Universal Robots PolyScope program: Sub_Centrifuge_V3.urp

Program Sub_Centrifuge_V3 (installation=default directory=/programs/03 Sub Routines createdIn=5.13.0 lastSavedIn=5.16.0 robotSerialNumber=20245590049)
Calibrated DH parameters: a=[0.000139, -0.197451, -0.383992, -0.000109, 0.000038, 0]; d=[0.162494, 274.063354, -251.846761, -22.083037, 0.099612, 0.099364]; alpha=[1.570089, 0.001374, 0.003592, 1.570222, -1.570187, 0]; deltaTheta=[0, 1.08787, 5.400214, -0.204909, 0.000001, 0]
InitVariablesNode variables(variable(name=DEV_CEN_PosRtr, expression=0))
BeforeStart
  Centrifuge := rpc_factory("xmlrpc","http://192.168.12.125:50002")
  Action :=  (valueSource=Operator message=What to do? valueType=Integer)
Robot Program (runOnlyOnce=true)
  Folder Handling
    SuppressedNode
      Folder PreSettings
        Folder Init Move Definitions [hidden by the author, left out]
        Folder Jig Definition [hidden by the author, left out]
        Folder Frame Definition [hidden by the author, left out]
        Folder Pose Definition [hidden by the author, left out]
    '===================='
    Switch expression=Action
      Case (caseValue=5)
        Folder Open
          Script: Centrifuge.open_hatch()
      Case (caseValue=6)
        Folder Close
          Script: Centrifuge.close_hatch()
      Case (caseValue=7)
        Folder Load
          DEV_CEN_CmdRslt := Centrifuge.move_rotor(DEV_CEN_PosRtr)
          If JNT_S≠[0,0,0,0,0,0]
            MoveJ speed 90 deg/s, acceleration 80 deg/s^2 (useActiveTCP=true positionType=JointAngles) feature=Base
              Waypoint Variable (Variable): motionParameters(blendRadius=0.05); variable=JNT_S
          MoveJ speed 90 deg/s, acceleration 80 deg/s^2 (useActiveTCP=true) feature=FRM_Reference
            If PSE_A_H≠p[0,0,0,0,0,0]
              Waypoint Variable (Variable): motionParameters(blendRadius=0.02); variable=PSE_A_H
            Waypoint Variable (Variable): variable=PSE_A
          If Centrifuge.posreached(DEV_CEN_PosRtr)
            MoveL speed 300 mm/s, acceleration 1200 mm/s^2 (useActiveTCP=true) feature=FRM_Reference
              If PSE_T_H≠p[0,0,0,0,0,0]
                Waypoint Variable (Variable): variable=PSE_T_H
              Waypoint Variable (Variable): motionParameters(jointSpeed=1.047198 jointAcceleration=1.396263 cartesianSpeed=0.075 cartesianAcceleration=1.2); variable=PSE_T
                Until TOOL_CONTACT_DETECTION (allowActions=true retraction=0.001 decelerationAcceleration=0.5 decelerationAngularAcceleration=34.906585)
                  Folder EOAT
                    URCap Gripper (Robotiq_Grippers, Robotiq Inc.) dataModel(position=88.72549019607843, force=25.0, speed=50.0, positionInDouble=88.72549019607843, forceInDouble=25.0, speedInDouble=50.0, slaveIds=[9], blocking=true)
                  Force Frame feature=Joint_6_name; selection=[0, 0, 0, 0, 0, 1]; wrench=[0, 0, 0, 0, 0, 0]; limitsForce=[0.15, 0.15, 0.15, 1.047198, 1.047198, 3.141593]; limitsMotion=[0.1, 0.1, 0.1, 0.349066, 0.349066, 0.349066]
                    Waypoint Variable (Variable): motionParameters(jointSpeed=1.047198 jointAcceleration=1.396263 cartesianSpeed=0.01 cartesianAcceleration=1.2); variable=PSE_T
              Folder EOAT
                URCap Gripper (Robotiq_Grippers, Robotiq Inc.) dataModel(position=70.09803921568627, force=50.0, speed=50.0, positionInDouble=70.09803921568627, forceInDouble=50.0, speedInDouble=50.0, slaveIds=[9], blocking=true)
              If PSE_R_H≠p[0,0,0,0,0,0]
                Waypoint Variable (Variable): motionParameters(blendRadius=0.01); variable=PSE_R
                Waypoint Variable (Variable): variable=PSE_R_H
              Else 
                Waypoint Variable (Variable): variable=PSE_R
      Case (caseValue=8)
        Folder Unload
          DEV_CEN_CmdRslt := Centrifuge.move_rotor(DEV_CEN_PosRtr)
          If JNT_S≠[0,0,0,0,0,0]
            MoveJ speed 90 deg/s, acceleration 80 deg/s^2 (useActiveTCP=true positionType=JointAngles) feature=Base
              Waypoint Variable (Variable): motionParameters(blendRadius=0.05); variable=JNT_S
          MoveJ speed 90 deg/s, acceleration 80 deg/s^2 (useActiveTCP=true) feature=FRM_Reference
            If PSE_A_H≠p[0,0,0,0,0,0]
              Waypoint Variable (Variable): motionParameters(blendRadius=0.02); variable=PSE_A_H
            Waypoint Variable (Variable): variable=PSE_A
          Folder EOAT
            URCap Gripper (Robotiq_Grippers, Robotiq Inc.) dataModel(position=70.09803921568627, force=50.0, speed=50.0, positionInDouble=70.09803921568627, forceInDouble=50.0, speedInDouble=50.0, slaveIds=[9], blocking=true)
          If Centrifuge.posreached(DEV_CEN_PosRtr)
            MoveL speed 300 mm/s, acceleration 1200 mm/s^2 (useActiveTCP=true) feature=FRM_Reference
              Waypoint Variable (Variable): motionParameters(jointSpeed=1.047198 jointAcceleration=1.396263 cartesianSpeed=0.1 cartesianAcceleration=1.2); variable=PSE_T
              Folder EOAT
                URCap Gripper (Robotiq_Grippers, Robotiq Inc.) dataModel(position=100.0, force=50.0, speed=50.0, positionInDouble=100.0, forceInDouble=50.0, speedInDouble=50.0, slaveIds=[9], blocking=true)
              If PSE_R_H≠p[0,0,0,0,0,0]
                Waypoint Variable (Variable): motionParameters(blendRadius=0.01); variable=PSE_R
                Waypoint Variable (Variable): variable=PSE_R_H
              Else 
                Waypoint Variable (Variable): variable=PSE_R
      Case (caseValue=9)
        Folder Start
          Script: Centrifuge.start()
      Case (caseValue=10)
        Folder Stop
          Script: Centrifuge.stop()
    '===================='
    Folder PostSettings [hidden by the author, left out]
